// TIA Portal V20 export
DATA_BLOCK "POS3_0_Antriebe_DB"   // DB24
// stored: AssignedProDiagFB POS3_0_Prodiag, InstanceOfName POS3_0_Antriebe, InstanceOfType FB
"POS3_0_Antriebe"
   // VAR
   //    "-1001T1_OM_PRM_Access_Instance" { S7_SetPoint := 'True'} : "OM_PRM_Access";
   //    "-1001T1_Oriental" { S7_SetPoint := 'True'} : "Oriental_AZD-KPN_Profinet";
   //    "-1002T2_OM_PRM_Access_Instance" { S7_SetPoint := 'True'} : "OM_PRM_Access";
   //    "-1002T2_Oriental_Drehachse" { S7_SetPoint := 'True'} : "Oriental_AZD-KPN_Profinet";
   //    Pos_Alt { S7_SetPoint := 'True'} : Real;
   //    Delta : Real;
   // END_VAR
BEGIN
END_DATA_BLOCK
